// TIA Portal V20 export
// export: Created 2026-11-12T11:17:33.7398542Z, ExportSetting WithDefaults, DisplayName Totally Integrated Automation Portal, DisplayVersion V20, DisplayName TIA Portal Openness, DisplayVersion V20, DisplayName TIA Portal Teamcenter Gateway, DisplayVersion V20, DisplayName TIA Portal Version Control Interface, DisplayVersion V20, DisplayName STEP 7 Professional, DisplayVersion V20, DisplayName STEP 7 CFC, DisplayVersion V20, DisplayName STEP 7 Safety, DisplayVersion V20, DisplayName WinCC Basic/Comfort/Advanced, DisplayVersion V20, DisplayName SIMATIC Visualization Architect, DisplayVersion V20, DisplayName WinCC Professional, DisplayVersion V20, DisplayName SIMATIC Visualization Architect, DisplayVersion V20, DisplayName WinCC Unified, DisplayVersion V20, DisplayName SIMATIC Visualization Architect, DisplayVersion V20
DATA_BLOCK "DB_Estacion"   // DB2
{ S7_Optimized_Access := 'TRUE' }
VERSION : 0.1
// stored: AutoNumber true, DBAccessibleFromOPCUA true, DBAccessibleFromWebserver true, IsOnlyStoredInLoadMemory false, IsRetainMemResEnabled false, IsWriteProtectedInAS false, MemoryReserve 100
   VAR
      Imagen_palet : Array[0..27] of Byte;
      App_inicio : Bool;
      App_en_reposo : Bool;
      App_terminada : Bool;
      App_alarma : Bool;
      App_rearme_requerido : Bool;
      Inhibir_cinta : Bool;
      Emergencia : Bool;
      Rearme : Bool;
   END_VAR
BEGIN
END_DATA_BLOCK
